(* IEC 61131-3 sources: SortJet_MasterSPS_Aufbau.fbsproj/Device.device.xml.v3^/Plc Logic.plclogic.xml.v3^/Application.application.xml.v3^/09_Station/Stationen/Aufgabe- Anlege- Wand[208]/0_Konfig, 3 files *)

(* ---- Antriebsinformationen_208.gvl ---- *)
(* METADATA
{
	"v3Meta": {
		"objectGuid": "0ee05288-750e-42b2-bc5b-835c7c5d3b07"
	}
}
*)
{attribute 'allow_unqualified_access'}
NAMESPACE Antriebsinformationen_208
VAR_GLOBAL

//-------------------------------------------------------------------------------------------------
// ANTRIEBSINFORMATION
//-------------------------------------------------------------------------------------------------

  apgInfoStation208Glastransport : ARRAY[cWAND_1..cANZAHL_WAENDE] OF AntriebsInformationen := [
    (
      wAchsID                                 :=     15,   // Achs ID aus dem EConSet
      stTyp                                   := 'Belt',  // Typ
      wpSchaltschrank                         :=   2080,  // Daten aus dem Schaltplan
      wpSchaltplanreihe                       :=      2,  // Daten aus dem Schaltplan
      wpSchaltplanseite                       :=    100,  // Daten aus dem Schaltplan
      rpMaxGeschwindigkeit                    :=   1000,  // [mm/s]   Max- Geschwindigkeit für den Automatikbetrieb
      rpHandGeschwindigkeit                   :=    333,  // [mm/s]   Hand- Geschwindigkeit
      rpReduzierteGeschwindigkeit             :=    250,  // [mm/s]   Reduzierte Geschwindigkeit
      rpReferenzGeschwindigkeit               :=     50,  // [mm/s]   Geschwindigkeit für die Referenzfahrt
      rpEinrichtGeschwindigkeit               :=    100,  // [mm/s]   Max Geschwindigkeit während der Einrichtung der Anlage
      rpMaxBeschleunigung                     :=   1500,  // [mm/s^2] Max Beschleunigung
      rpMaxVerzoegerung                       :=   1500,  // [mm/s^2] Max Verzoegerung
      rpMaxRuckzeit                           :=    100,  // [ms]     Ruckzeit des Antriebs
      rpReduzierteBeschleunigung              :=    500,  // [mm/s^2] Reduzierte Beschleunigung
      rpReduzierteVerzoegerung                :=    500,  // [mm/s^2] Reduzierte Verzoegerung
      rpBeschleunigungFremdanlage             :=   1000,  // [mm/s^2] Beschleunigung zu einer Fremdanlage
      rpGeschwindigkeitMessen                 :=    667,  // [mm/s] Geschwindigkeit beim Scheiben messen
      rpGeschwindigkeitSystemcheck            :=  500.0,  // [mm/s]   Geschwindigkeit im Systemcheck (nur Glastransport)
      rpGeschwindigkeitSystemcheckReduzierung :=  167.0,  // [mm/s]   Geschwindigkeit im Systemcheck bei belegtem Vorstop-Sensor (nur Glastransport)
      stOptionen                              := ( eEndschalterQuelle    := Endschalterquelle_EN.KEINE,     // Hardware-Endschalter: KEINE, UMRICHTER oder SPS
                                                   bVersorgungUeberXVR   := FALSE,                          // XVR-Modus: brueckt Hauptschalter 400 V und LS 230 V
                                                   bBremseLoesenFreigabe := FALSE )                         // Der Antrieb darf über eine Betriebsart die Bremse lösen
    )];

  apgInfoStation208GlastransportSlave : ARRAY[cWAND_1..cANZAHL_WAENDE] OF AntriebsInformationen := [
    (
      wAchsID                                 :=     65,   // Achs ID aus dem EConSet
      stTyp                                   := 'Belt',  // Typ
      wpSchaltschrank                         :=   2080,  // Daten aus dem Schaltplan
      wpSchaltplanreihe                       :=      2,  // Daten aus dem Schaltplan
      wpSchaltplanseite                       :=    100,  // Daten aus dem Schaltplan
      rpMaxGeschwindigkeit                    :=   1000,  // [mm/s]   Max- Geschwindigkeit für den Automatikbetrieb
      rpHandGeschwindigkeit                   :=    333,  // [mm/s]   Hand- Geschwindigkeit
      rpReduzierteGeschwindigkeit             :=    250,  // [mm/s]   Reduzierte Geschwindigkeit
      rpReferenzGeschwindigkeit               :=     50,  // [mm/s]   Geschwindigkeit für die Referenzfahrt
      rpEinrichtGeschwindigkeit               :=    100,  // [mm/s]   Max Geschwindigkeit während der Einrichtung der Anlage
      rpMaxBeschleunigung                     :=   1500,  // [mm/s^2] Max Beschleunigung
      rpMaxVerzoegerung                       :=   1500,  // [mm/s^2] Max Verzoegerung
      rpMaxRuckzeit                           :=    100,  // [ms]     Ruckzeit des Antriebs
      rpReduzierteBeschleunigung              :=    500,  // [mm/s^2] Reduzierte Beschleunigung
      rpReduzierteVerzoegerung                :=    500,  // [mm/s^2] Reduzierte Verzoegerung
      rpBeschleunigungFremdanlage             :=   1000,  // [mm/s^2] Beschleunigung zu einer Fremdanlage
      rpGeschwindigkeitMessen                 :=    667,  // [mm/s] Geschwindigkeit beim Scheiben messen
      rpGeschwindigkeitSystemcheck            :=  500.0,  // [mm/s]   Geschwindigkeit im Systemcheck (nur Glastransport)
      rpGeschwindigkeitSystemcheckReduzierung :=  167.0,  // [mm/s]   Geschwindigkeit im Systemcheck bei belegtem Vorstop-Sensor (nur Glastransport)
      stOptionen                              := ( eEndschalterQuelle    := Endschalterquelle_EN.KEINE,     // Hardware-Endschalter: KEINE, UMRICHTER oder SPS
                                                   bVersorgungUeberXVR   := FALSE,                          // XVR-Modus: brueckt Hauptschalter 400 V und LS 230 V
                                                   bBremseLoesenFreigabe := FALSE )                         // Der Antrieb darf über eine Betriebsart die Bremse lösen
    )];

  apgInfoStation208Messachse :  AntriebsInformationen :=
    (
      wAchsID                                 :=        16,   // Achs ID aus dem EConSet
      stTyp                                   := 'Measure',  // Typ
      wpSchaltschrank                         :=      2081,  // Daten aus dem Schaltplan
      wpSchaltplanreihe                       :=         2,  // Daten aus dem Schaltplan
      wpSchaltplanseite                       :=       100,  // Daten aus dem Schaltplan
      rpMaxGeschwindigkeit                    :=      1000,  // [mm/s]   Max- Geschwindigkeit für den Automatikbetrieb
      rpHandGeschwindigkeit                   :=       333,  // [mm/s]   Hand- Geschwindigkeit
      rpReduzierteGeschwindigkeit             :=         0,  // [mm/s]   Reduzierte Geschwindigkeit
      rpReferenzGeschwindigkeit               :=        50,  // [mm/s]   Geschwindigkeit für die Referenzfahrt
      rpEinrichtGeschwindigkeit               :=         0,  // [mm/s]   Max Geschwindigkeit während der Einrichtung der Anlage
      rpMaxBeschleunigung                     :=      2500,  // [mm/s^2] Max Beschleunigung
      rpMaxVerzoegerung                       :=      2500,  // [mm/s^2] Max Verzoegerung
      rpMaxRuckzeit                           :=       500,  // [ms]     Ruckzeit des Antriebs
      rpReduzierteBeschleunigung              :=       500,  // [mm/s^2] Reduzierte Beschleunigung
      rpReduzierteVerzoegerung                :=       500,  // [mm/s^2] Reduzierte Verzoegerung
      rpBeschleunigungFremdanlage             :=         0,  // [mm/s^2] Beschleunigung zu einer Fremdanlage
      rpGeschwindigkeitMessen                 :=         0,  // [mm/s] Geschwindigkeit beim Scheiben messen
      rpGeschwindigkeitSystemcheck            :=     500.0,  // [mm/s]   Geschwindigkeit im Systemcheck (nur Glastransport)
      rpGeschwindigkeitSystemcheckReduzierung :=     167.0,  // [mm/s]   Geschwindigkeit im Systemcheck bei belegtem Vorstop-Sensor (nur Glastransport)
      stOptionen                              := ( eEndschalterQuelle    := Endschalterquelle_EN.UMRICHTER, // Hardware-Endschalter: KEINE, UMRICHTER oder SPS
                                                   bVersorgungUeberXVR   := FALSE,                          // XVR-Modus: brueckt Hauptschalter 400 V und LS 230 V
                                                   bBremseLoesenFreigabe := FALSE )                         // Der Antrieb darf über eine Betriebsart die Bremse lösen
    );

  apgInfoStation208Kippen : AntriebsInformationen :=
    (
      wAchsID                                 :=     65,  // Achs ID aus dem EConSet
      stTyp                                   := 'Tilt',  // Typ
      wpSchaltschrank                         :=      0,  // Daten aus dem Schaltplan
      wpSchaltplanreihe                       :=     02,  // Daten aus dem Schaltplan
      wpSchaltplanseite                       :=      0,  // Daten aus dem Schaltplan
      rpMaxGeschwindigkeit                    :=      0,  // [Grad/s]   Max- Geschwindigkeit für den Automatikbetrieb
      rpHandGeschwindigkeit                   :=      0,  // [Grad/s]   Hand- Geschwindigkeit
      rpReduzierteGeschwindigkeit             :=      0,  // [Grad/s]   Reduzierte Geschwindigkeit
      rpReferenzGeschwindigkeit               :=      0,  // [Grad/s]   Geschwindigkeit für die Referenzfahrt
      rpEinrichtGeschwindigkeit               :=      0,  // [Grad/s]   Max Geschwindigkeit während der Einrichtung der Anlage
      rpMaxBeschleunigung                     :=      0,  // [Grad/s^2] Max Beschleunigung
      rpMaxVerzoegerung                       :=      0,  // [Grad/s^2] Max Verzoegerung
      rpMaxRuckzeit                           :=      0,  // [ms] Ruckzeit des Antriebs
      rpReduzierteBeschleunigung              :=      0,  // [Grad/s^2] Reduzierte Beschleunigung
      rpReduzierteVerzoegerung                :=      0,  // [Grad/s^2] Reduzierte Verzoegerung
      rpBeschleunigungFremdanlage             :=      0,  // [Grad/s^2] Beschleunigung zu einer Fremdanlage
      rpGeschwindigkeitMessen                 :=      0,  // [Grad/s] Geschwindigkeit beim Scheiben messen
      rpGeschwindigkeitSystemcheck            :=  500.0,  // [mm/s]   Geschwindigkeit im Systemcheck (nur Glastransport)
      rpGeschwindigkeitSystemcheckReduzierung :=  167.0,  // [mm/s]   Geschwindigkeit im Systemcheck bei belegtem Vorstop-Sensor (nur Glastransport)
      stOptionen                              := ( eEndschalterQuelle    := Endschalterquelle_EN.KEINE,     // Hardware-Endschalter: KEINE, UMRICHTER oder SPS
                                                   bVersorgungUeberXVR   := FALSE,                          // XVR-Modus: brueckt Hauptschalter 400 V und LS 230 V
                                                   bBremseLoesenFreigabe := FALSE )                         // Der Antrieb darf über eine Betriebsart die Bremse lösen
    );

END_VAR

END_NAMESPACE

(* ---- MK_Station_208.gvl ---- *)
(* METADATA
{
	"v3Meta": {
		"objectGuid": "8432a7e6-a09e-4ecf-ad2f-9f4275e97011"
	}
}
*)
{attribute 'allow_unqualified_access'}
NAMESPACE MK_Station_208
VAR_GLOBAL

//-------------------------------------------------------------------------------------------------
// MASCHINEPARAMETER: ANLEGE- ABNAHME- WAND
//-------------------------------------------------------------------------------------------------

  apgMKStation208 : Parameter_Station :=
    (
      stStationsNummern                     := ( NummerIntern :=  208,                                                       // Stationsnummer fuer das MMI und die Stationsangabe der Meldungen
                                                 NummerExtern := 1208,                                                       // Stationsnummer fuer Bedienermeldungen
                                                 NummerSPS    :=  208                                                        // Stationsnummer SPS-intern (Indizes)
                                               ),
      bDeaktivieren                         := FALSE,                                                                        // Station deaktiviert (keine Auftraege, keine Referenzfahrt)
      wMeldungsNummer                       := 1830,                                                                         // Basis-Meldungsnummer (WatchIO)
      eStationsTyp                          := eStation,                                                                     // Typ der Station
      eaAutomatikkreis                      := [eAutomatikkreis_1],                                                          // Automatikkreise, zu denen die Station gehoert
      eaSicherheitskreis                    := [eSicherheitskreis_Undefiniert],                                              // Sicherheitskreise, in die die Station eingebunden ist
      // astSicherheitskreisTeilabschaltung
      eSystemcheckZyklus                    := eSystemcheckZyklus_1,                                                         // In welchem Zyklus des Systemchecks die Station geprueft wird
      stSchnittstellendaten                 := ( wVorgaengerStation := cSTATION_DEFAULT,                                     // Station vor dieser Station (cSTATION_DYNAMISCH bei mehreren)
                                                 wNachfolgerStation := cSTATION_207,                                         // Station nach dieser Station (cSTATION_DYNAMISCH bei mehreren)
                                                 bStationIstShuttle := FALSE                                                 // Station ist ein Shuttle
                                               ),
      stStationsOptionen                    := ( stSystemcheck :=  ( bScheibenVermessenSystemCheck               := FALSE,   // Scheiben im Systemcheck vermessen
                                                                     bScheibeNachSystemcheckAufAuslauf           := TRUE,    // Scheibe nach dem Systemcheck auf den Auslaufsensor fahren
                                                                     bSystemCheckMitVorgaengerBatchTransport     := FALSE,   // derzeit ohne Funktion
                                                                     bSystemCheckMitNachfolgerBatchTransport     := FALSE,   // derzeit ohne Funktion
                                                                     bOptionSystemCheckScheibeMittigLegen        := FALSE ), // derzeit ohne Funktion

                                                 // stTransfershuttle
                                                 stGlastransport :=  ( bVortransport                             := FALSE,   // Vortransport aktivieren [Bsp.: Nach einem Eintransport mit gesetztem Bit <Letzte Scheibe>]
                                                                       bTransportMasterSlaveEintransport         := FALSE,   // derzeit ohne Funktion
                                                                       bTransportMasterSlaveAustransport         := TRUE ,   // Austransport als Slave auf die Achse des Nachfolgers
                                                                       bGLasUebernahmeSenkrecht                  := FALSE,   // RKT - Eintransport in Senkrechter-Position bzw. in Waagerechter- Position [default]
                                                                       bAustransportISOLinie                     := FALSE,   // Austransport an eine ISO-Linie
                                                                       bScheibenVermessen                        := TRUE,    // Scheibenmessung am Anlegetisch/Anlegewand
                                                                       bMessrichtungNegativ                      := FALSE,   // Negative Fahrtrichtung beim Messen
                                                                       bScheibenmessungEintransport              := FALSE,   // Scheibenmessung beim Eintransport
                                                                       bScheibenmessungSensorVorabAuslauf        := TRUE     // Scheibenmessung mit SensorVorabAuslauf z.B. Anlegewand
                                                                      ),
                                                 stAnlegetisch   :=  ( bIstAnlegestation                         := TRUE,    // Station an der Scheiben angelegt werden [Anlegetisch, Anlegewand]; im Systemcheck-Verbund nur mit genau einer Scheibe
                                                                       bAnschlagAutomatischAusfahren             := FALSE,   // Anschlaege beim Anlegen automatisch ausfahren (Vorgabe, am Taster umschaltbar)
                                                                       bAnlegetischMitEintransportVorgaenger     := FALSE    // VSG: Station entscheidet selbst zwischen Eintransport vom Vorgaenger und Anlegen
                                                                      ),
                                                 // stEckuebergabe
                                                 // stDrehstation
                                                 bVorAbKomponentenAnsteuerung              := FALSE,                         // VorAbKomponentenAnsteuerung Auftraege werden bearbeitet
                                                 bVerstellungEinAusGefahrenLogikDrehen     := FALSE,                         // Verstellung: Logik ein-/ausgefahren gedreht
                                                 bLangsamfahrtNockenQuerfahrtAktivieren    := FALSE,                         // Querfahrt: Langsamfahrt-Nocken auswerten
                                                 bSKBlockierenDurchVorabSensoren           := FALSE,                         // Vorab-Sensoren belegt blockieren das Oeffnen des Sicherheitskreises
                                                 bStationLeerfahrenBeiSkAnforderung        := FALSE,                         // Station bei Anforderung Sicherheitskreis leerfahren
                                                 bScheibeAbnehmenNachEintransport          := TRUE,                          // Scheibe nach dem Eintransport wieder abnehmen
                                                 bGlasAbgenommenAutomatischQuittieren      := FALSE                          // derzeit ohne Funktion
                                               ),
      stStationsAufbau                      := ( bGeblase                      := [ cANZAHL_WAENDE(FALSE) ],                 // Ausbaustufe: Geblaese je Wand
                                                 bGlastransport                := [ TRUE ],                                  // Ausbaustufe: Glastransport je Wand
                                                 bKippen                       := [ cANZAHL_WAENDE(FALSE) ],                 // Ausbaustufe: Kippen je Wand
                                                 bKippenSchuetz                := FALSE,                                     // Kippen ueber Schuetz statt Umrichter
                                                 bTransportVerstellung         := [ cANZAHL_WAENDE(FALSE) ],                 // Ausbaustufe Shuttle: Transport-/Dickenverstellung je Wand
                                                 bHub                          := FALSE,                                     // Ausbaustufe: Hub der Station
                                                 bHubrahmen                    := FALSE,                                     // Ausbaustufe: Hubrahmen (Riemen heben/senken)
                                                 bDrehen                       := FALSE,                                     // Ausbaustufe: Drehen
                                                 bQuerachse                    := FALSE,                                     // Ausbaustufe: Querachse
                                                 bMessachse                    := TRUE,                                      // Ausbaustufe: Messachse (Anlegetisch, Anlegewand)
                                                 bDruckluft                    := FALSE,                                     // Druckluftueberwachung vorhanden
                                                 bAnschlag                     := FALSE,                                     // Ausbaustufe: Ausrichtanschlaege
                                                 bSensorAuslauf                := TRUE,                                      // Auslaufsensor vorhanden
                                                 bSensorEinlauf                := TRUE,                                      // Einlaufsensor vorhanden
                                                 bSensorEinlaufStopp           := FALSE,                                     // Shuttle: zusaetzlicher Stopp-Sensor am Einlauf (ohne: Einlaufsensor), Gegenstueck zum Auslauf-Stopp im Rueckwaertstransport
                                                 bSensorAuslaufStopp           := FALSE,                                     // Shuttle: zusaetzlicher Stopp-Sensor am Auslauf (ohne: Auslaufsensor), Verfahrfreigabe und Scheibe hat Shuttle verlassen
                                                 bDurchlaufSperreZumNachfolger := TRUE,                                      // Ausbaustufe: bewegliche Abschrankung zum Nachfolger
                                                 bQuerfahrt                    := FALSE,                                     // Ausbaustufe: Querfahrt
                                                 bWandverstellung              := [ FALSE ],                                 // Ausbaustufe Station: Wandverstellung je Wand
                                                 bWandverstellungMotorisch     := FALSE,                                     // Shuttle: Transport-/Wandverstellung mit Antrieb statt pneumatisch
                                                 bRoellchenleiste              := [ FALSE ],                                 // Ausbaustufe Station: Roellchenleiste je Wand
                                                 bDurchgang                    := FALSE,                                     // Station ist Teil eines Durchgangs (belegt = Oeffnen blockiert)
                                                 bSlaveAntrieb                 := FALSE,                                     // Glastransport mit Slave-Antrieb
                                                 bRolltor                      := FALSE,                                     // Ausbaustufe Faecherwagen: Rolltor
                                                 bKlemmzylinder                := FALSE,                                     // Ausbaustufe Faecherwagen: Klemmzylinder fixiert den Oberrahmen beim Ein- und Ausschleusen
                                                 bGreifer                      := [cANZAHL_WAENDE(FALSE)],                   // Shuttle: Greifer je Wand (Scheibe aus dem Faecherwagen ziehen bzw. hineinschieben)
                                                 bRFID                         := FALSE,                                     // RFID-Leser vorhanden
                                                 bAGV                          := FALSE,                                     // Ausbaustufe Faecherwagen: Betrieb mit AGV
                                                 bKipparme                     := FALSE,                                     // Ausbaustufe: Kipparme
                                                 bMessachseAmEndeVomTisch      := FALSE,                                     // Messachse am Ende des Tisches (Hoehenfehler fragt den Bediener)
                                                 bDLSSchmiersystem             := FALSE,                                     // Zentralschmierung DLS vorhanden
                                                 bGlastransportSlaveVorhanden  := FALSE,                                     // Glastransport mit Slave-Antrieb (Meldungen/Ueberwachung Slave)
                                                 wHydraulikstation             := 0                                          // Faecherwagen Hydraulik: zugeordnete Hydraulikstation (cHYDRAULIKSTATION_x), 0 = keine
                                               ),
      stStationsParameter                   := ( rLaengeUebergroesseScheibe              := 6000,                            // Shuttle: ab dieser Scheibenlaenge gilt die Scheibe als uebergross [mm]
                                                 rMinGlasHoeheAutomatischenEintransport  := 0.0,                             // VSG: Mindesthoehe fuer automatischen Eintransport [mm]
                                                 rMinGlasLaengeAutomatischenEintransport := 0.0,                             // VSG: Mindestlaenge fuer automatischen Eintransport [mm]
                                                 wMaximaleAnzahlAktiverAuftraege         := 0,                               // derzeit ohne Funktion
                                                 rMinPosSwEsEingrenzung                  := 0.0,                             // Externer zusaetzlicher Software-Endschalter MIN; 0 = inaktiv; darf den MK-MIN nur weiter eingrenzen
                                                 rMaxPosSwEsEingrenzung                  := 0.0,                             // Externer zusaetzlicher Software-Endschalter MAX; 0 = inaktiv; darf den MK-MAX nur weiter eingrenzen
                                                 rPosFreigabePufferAusfahren             := 0.0                              // derzeit ohne Funktion
                                               ),
      // stFremdanlage
      stGlasdaten                           := [( rlMinGlasLaenge := 350,                                                    // minimal zulässige GlasLänge
                                                  rlMaxGlasLaenge := 2500,                                                   // maximale zulässige GlasLänge
                                                  rlMinGlasHoehe  := 190,                                                    // minimal zulässige GlasHöhe
                                                  rlMaxGlasHoehe  := 1800,                                                   // maximale zulässige GlasHöhe
                                                  rlMinGlasDicke  := 3,                                                    // minimal zulässige GlasDicke
                                                  rlMaxGlasDicke  := 12.76,                                                     // maximal zulaessige Glasdicke [mm]
                                                  rlLaengeMaxGlas := 0.0                                                     // maximal zulaessige Glaslaenge [mm]
                                               )]
      // astShuttleAnhaltenQuellen
     );

   apgMKStation208Glastransport : ARRAY[cWAND_1..cANZAHL_WAENDE] OF Parameter_Glastransport := [
    (
      rLaengeStation                        :=  3300, // Länge der Station
      rScheibenabstand                      :=   300, // Der Abstand zwischen zwei Scheiben auf der Station
      rWegUeberAuslauf                      :=    50, // Weg ueber den Auslaufsensor hinaus [mm]
      rWegUeberEinlauf                      :=    50, // Weg ueber den Einlaufsensor hinaus [mm]
      rWegUeberSensorenSystemCheck          :=    15, // Der Weg der Ueber ein die Sensoren zum vermessen der Scheiben
      rUeberwachungAuslaufsensor            :=   500, // Ueberwachung des Auslaufsensors [Strecke in der der Auslaufsensor Frei / ueberfahren werden soll]
      rUeberwachungEinlaufsensor            :=   500, // Ueberwachung des Einlaufsensors [Strecke in der der Einlaufsensor Frei / ueberfahren werden soll]
      rWegUeberEinlaufEintransport          :=    30, // Eintransport vorwaerts: Abstand Scheibenhinterkante zum Einlaufsensor [mm]
      rWegUeberEinlaufAustransport          :=    30, // Lage Auf Einlauf: Scheibe liegt um diesen Weg auf dem Einlaufsensor [mm]
      rWegUeberAuslaufEintransport          :=    30, // Eintransport rueckwaerts: Abstand Scheibenhinterkante zum Auslaufsensor [mm]
      rWegUeberAuslaufAustransport          :=    15, // Lage Auf Auslauf: Weg ueber den Auslaufsensor hinaus [mm]
      rWegEinlaufsensorZuVorStopSensor      :=  3160, // Beschreibt den Weg vum eine Scheibe beim EIntransport vom Einlaufsensor bis ueberden Vorabstopsensor zu verfahren
      rMesstoleranz                         :=    10, // Toleranz-Mass fuer die Scheibenlaengenmessung
      rMessstrecke                          :=  2904, // Beschreibt die Strecke ziwischen 2 Sensoren die der Antrieb verfaehrt
      rWegstreckeBisZurVerzoegerung         :=  2660  // Beschreibt die Strecke die gefahren werden soll bis der Antrieb abgebremst werden soll, dies gilt fuer Eintransportauftraege die das Bit "Letzte Scheibe" gesetzt haben
    )];

  apgMKStation208Messachse: Parameter_Messachse :=
    (
      rKorrekturOffset                      :=    0, // Korrektur der Position um einen Bestimmten Wert (Offset)
      rStreckePositionieren                 :=    0, // ?
      rPositionUeberScheibenhoehe           := 0.0,  // Position der Zentrierleiste ueber dem Glas so dass das Glas angelegt werden kann
      rVerfahrbereichsOffset                := 0.0,  // Korrektur des Verfahrens wenn
      rKorrekturOffsetVSGEintransport       := 0.0,  // Korrektur der Position um einen Bestimmten Wert (Offset) beim Eintransport von VSG
      rOffsetMessung                        := 0.0,  // ?
      rToleranz                             := 0.0,  // Toleranzwert in der Ausmessung der Höhe
      rAbstandSensorenOberUndUnterkante     := 0.0,  // Rechnerischer Abstand zwischen dem Sensor der die Scheibenunterkante misst und dem Sensor der die Scheibenoberkante misst
      rOffsetNullLinie                      := 0.0   // Offset das auf den Wert des Abstands zur Null-Linie aufgerechnet wird, um dies evtl zu korrigieren
    );

  apgMKStation208Kippen : ARRAY[cWAND_1..cANZAHL_WAENDE] OF Parameter_Kippen := [
    (
      tZeitlicheUeberwachungKippen          := TIME#5000MS, // [ms \ s] Verwendet fuer Antriebe die Ueber einen Schuetz angesteuert werden
      tZeitAntriebsfreigabeErhalten         :=  TIME#180S,  // [ms \ s] Energieeinsparrung: Zeiteinheit nach der die Antriebsfreigabe entzogen werden soll wenn keine Aktion ansteht [1 s = 1000 ms ]
      rToleranz                             :=          1,  // Toleranz beim Entscheiden der aktuellen Position
      rPosition0Grad                        :=          0,  // Waagerechte- Position 0 Grad: Position auf die die Station gehoben werden soll
      rPosition90Grad                       :=          0,  // Senkrechte-Position 90 Grad : Position auf die die Station gesenkt werden soll
      bKippenMitSchuetz                     :=      FALSE,  // Kippen per Umrichter oder Schütz
      rPosition84Grad                       := 0.0,         // Senkrechte- Position 84 Grad: Position auf die die Station gehoben werden soll
      rPosition88_5Grad                     := 0.0,         // Senkrechte- Position 84 Grad: Position auf die die Station gehoben werden soll
      rPosition96Grad                       := 0.0          // Senkrechte-Position 96 Grad : Position auf die die Station gesenkt werden soll
    )];

END_VAR
END_NAMESPACE

(* ---- Konfiguration_208.gvl ---- *)
(* METADATA
{
	"v3Meta": {
		"objectGuid": "94633f29-785d-43e8-8fe9-544c355e9fea"
	}
}
*)
{attribute 'allow_unqualified_access'}
NAMESPACE Konfiguration_208
VAR_CONFIG

  // Taster
  Globale_Bausteine.Combiwand208.in_bFussTasterGlasAngelegt                               AT %MX1.0    : BOOL; // OPTION - Signal Scheibe ist angelegt Fusstaster
  Globale_Bausteine.Combiwand208.in_bTasterGlasAngelegt                                   AT %IX3.7    : BOOL; // IO-L - 208 quittieren Scheibe aufgelegt
  Globale_Bausteine.Combiwand208.in_bTasterFehlmessungQuittiern                           AT %IX4.0    : BOOL; // IO-L - 208 Fehlmessung quittieren
  Globale_Bausteine.Combiwand208.in_bKnebelGlastransportZurueck                           AT %IX4.2    : BOOL; // IO-L - 208 Riemen zurueck
  Globale_Bausteine.Combiwand208.in_bKnebelGlastransportVor                               AT %IX4.1    : BOOL; // IO-L - 208 Riemen vor
  Globale_Bausteine.Combiwand208.in_bTasterGlasbruch                                      AT %IX4.3    : BOOL; // IO-L - 208 Glasbruch
  Globale_Bausteine.Combiwand208.in_bTasterQuittierungGlasAbgenommen                      AT %IX3.7    : BOOL; // IO-L - 208 quittieren Scheibe aufgelegt (gleicher Taster wie Glas angelegt)

  // Lampen/Ampel
  Globale_Bausteine.Combiwand208.out_bAmpelSignalGruen                                    AT %QX5.0    : BOOL; // IO-L - 208 Freigabe Scheibe anlegen Ampel gruen
  Globale_Bausteine.Combiwand208.out_bSignalScheibeAufgegeben                             AT %QX4.5    : BOOL; // IO-L - 208 quittieren Scheibe aufgelegt
  Globale_Bausteine.Combiwand208.out_bSignalScheibeFehlmessung                            AT %QX4.6    : BOOL; // IO-L - 208 Scheibe Fehlmessung
  Globale_Bausteine.Combiwand208.out_bSignalScheibeGlasbruch                              AT %QX4.7    : BOOL; // IO-L - 208 Glasbruch Meldung
  Globale_Bausteine.Combiwand208.out_bSignalScheibeAbnehmen                               AT %MX2080.1 : BOOL; // OPTION

  // Bewegliche Abschrankung zum Nachfolger (geschlossen kommt ueber die Safety)
  Globale_Bausteine.Combiwand208.in_bSensorAbschrankungOffen                              AT %IX9.0    : BOOL; // IO-L - 208 bewegliche Abschrankung offen
  Globale_Bausteine.Combiwand208.out_bAbschrankungEinfahren                               AT %QX10.4   : BOOL; // IO-L - 208 bewegliche Abschrankung einfahren (oeffnen)
  Globale_Bausteine.Combiwand208.out_bAbschrankungAusfahren                               AT %QX10.5   : BOOL; // IO-L - 208 bewegliche Abschrankung ausfahren (schliessen)

  // Lichtschranke
  Globale_Bausteine.Combiwand208.in_bLichtschrankeQuittiert                               AT %MX1.1    : BOOL; // OPTION
  Globale_Bausteine.Combiwand208.in_bLichtschrankeFehler                                  AT %MX1.1    : BOOL; // OPTION
  Globale_Bausteine.Combiwand208.out_bLichtschrankeAusgeloest                             AT %MX2080.2 : BOOL; // OPTION - Lichtschranke an der Station ausgelöst und nicht quittiert

  // Gebläse
  Globale_Bausteine.Combiwand208.in_bTasterGeblaeseEin                                    AT %MX1.0     : BOOL; // OPTION - Taster Geblaese ein
  Globale_Bausteine.Combiwand208.in_bMotorschutzGeblaese_Ok                               AT %MX1.1     : BOOL; // OPTION - Motorschutzschalter / Sicherung des Antriebs
  Globale_Bausteine.Combiwand208.out_bGeblaeseEin                                         AT %MX2080.3  : BOOL; // OPTION - Geblaese starten (Schuetz)

  // Dickenverstellung
  Globale_Bausteine.Combiwand208.Dickenverstellung.in_bStatusZylinder1Ausgefahren         AT %MX1.0     : BOOL; // OPTION
  Globale_Bausteine.Combiwand208.Dickenverstellung.in_bStatusZylinder1Eingefahren         AT %MX1.0     : BOOL; // OPTION
  Globale_Bausteine.Combiwand208.Dickenverstellung.in_bStatusZylinder2Ausgefahren         AT %MX1.0     : BOOL; // OPTION
  Globale_Bausteine.Combiwand208.Dickenverstellung.in_bStatusZylinder2Eingefahren         AT %MX1.0     : BOOL; // OPTION

  Globale_Bausteine.Combiwand208.Dickenverstellung.out_bZylinder1Ausfahren                AT %MX2080.4  : BOOL; // OPTION
  Globale_Bausteine.Combiwand208.Dickenverstellung.out_bZylinder1Einfahren                AT %MX2080.5  : BOOL; // OPTION
  Globale_Bausteine.Combiwand208.Dickenverstellung.out_bZylinder2Ausfahren                AT %MX2080.6  : BOOL; // OPTION
  Globale_Bausteine.Combiwand208.Dickenverstellung.out_bZylinder2Einfahren                AT %MX2080.7  : BOOL; // OPTION

  // Kippen
  Globale_Bausteine.Combiwand208.Kippen.in_bMotorschutzschalter_OK                        AT %MX1.1     : BOOL; // OPTION
  Globale_Bausteine.Combiwand208.Kippen.in_bMotorstarter_OK                               AT %MX1.1     : BOOL; // OPTION
  Globale_Bausteine.Combiwand208.Kippen.in_bLSBremse_OK                                   AT %MX1.1     : BOOL; // OPTION
  Globale_Bausteine.Combiwand208.Kippen.in_bLS400V_OK                                     AT %MX1.1     : BOOL; // OPTION

  Globale_Bausteine.Combiwand208.Kippen.out_bKippen84Grad                                 AT %MX2081.0  : BOOL; // OPTION
  Globale_Bausteine.Combiwand208.Kippen.out_bKippen90Grad                                 AT %MX2081.1  : BOOL; // OPTION
  Globale_Bausteine.Combiwand208.Kippen.out_bBremseLoesen                                 AT %MX2081.2  : BOOL; // OPTION
  Globale_Bausteine.Combiwand208.Kippen.out_bReset                                        AT %MX2081.3  : BOOL; // OPTION

  // Nicht vorhandene Komponenten (der Basic erwartet sie, die Instanzen bleiben deaktiviert): Eingaenge auf %MX1.x, Ausgaenge auf freie Merker

  // Hub (unbenutzt)
  Globale_Bausteine.Combiwand208.HubUnbenutzt.in_bSensorNichtUnten                                AT %MX1.0   : BOOL; // OPTION
  Globale_Bausteine.Combiwand208.HubUnbenutzt.in_bSensorNichtOben                                 AT %MX1.0   : BOOL; // OPTION
  Globale_Bausteine.Combiwand208.HubUnbenutzt.in_bMotorstarter_OK                                 AT %MX1.1   : BOOL; // OPTION
  Globale_Bausteine.Combiwand208.HubUnbenutzt.in_bLSBremse_OK                                     AT %MX1.1   : BOOL; // OPTION
  Globale_Bausteine.Combiwand208.HubUnbenutzt.in_bLS400V_OK                                       AT %MX1.1   : BOOL; // OPTION
  Globale_Bausteine.Combiwand208.HubUnbenutzt.out_bHubAbSetzen                                    AT %MX2081.4 : BOOL; // OPTION
  Globale_Bausteine.Combiwand208.HubUnbenutzt.out_bHubAufSetzen                                   AT %MX2081.5 : BOOL; // OPTION
  Globale_Bausteine.Combiwand208.HubUnbenutzt.out_bReset                                          AT %MX2081.6 : BOOL; // OPTION
  Globale_Bausteine.Combiwand208.HubUnbenutzt.out_bBremseLoesen                                   AT %MX2081.7 : BOOL; // OPTION

  // Roellchenleiste (unbenutzt)
  Globale_Bausteine.Combiwand208.RoellchenleisteUnbenutzt.in_bStatusZylinder1Ausgefahren          AT %MX1.0   : BOOL; // OPTION
  Globale_Bausteine.Combiwand208.RoellchenleisteUnbenutzt.in_bStatusZylinder1Eingefahren          AT %MX1.0   : BOOL; // OPTION
  Globale_Bausteine.Combiwand208.RoellchenleisteUnbenutzt.in_bStatusZylinder2Ausgefahren          AT %MX1.0   : BOOL; // OPTION
  Globale_Bausteine.Combiwand208.RoellchenleisteUnbenutzt.in_bStatusZylinder2Eingefahren          AT %MX1.0   : BOOL; // OPTION
  Globale_Bausteine.Combiwand208.RoellchenleisteUnbenutzt.out_bZylinder1Ausfahren                 AT %MX2082.0 : BOOL; // OPTION
  Globale_Bausteine.Combiwand208.RoellchenleisteUnbenutzt.out_bZylinder1Einfahren                 AT %MX2082.1 : BOOL; // OPTION
  Globale_Bausteine.Combiwand208.RoellchenleisteUnbenutzt.out_bZylinder2Ausfahren                 AT %MX2082.2 : BOOL; // OPTION
  Globale_Bausteine.Combiwand208.RoellchenleisteUnbenutzt.out_bZylinder2Einfahren                 AT %MX2082.3 : BOOL; // OPTION

  // Wandverstellung (unbenutzt)
  Globale_Bausteine.Combiwand208.WandverstellungUnbenutzt.in_bStatusZylinder1Ausgefahren          AT %MX1.0   : BOOL; // OPTION
  Globale_Bausteine.Combiwand208.WandverstellungUnbenutzt.in_bStatusZylinder1Eingefahren          AT %MX1.0   : BOOL; // OPTION
  Globale_Bausteine.Combiwand208.WandverstellungUnbenutzt.in_bStatusZylinder2Ausgefahren          AT %MX1.0   : BOOL; // OPTION
  Globale_Bausteine.Combiwand208.WandverstellungUnbenutzt.in_bStatusZylinder2Eingefahren          AT %MX1.0   : BOOL; // OPTION
  Globale_Bausteine.Combiwand208.WandverstellungUnbenutzt.out_bZylinder1Ausfahren                 AT %MX2082.4 : BOOL; // OPTION
  Globale_Bausteine.Combiwand208.WandverstellungUnbenutzt.out_bZylinder1Einfahren                 AT %MX2082.5 : BOOL; // OPTION
  Globale_Bausteine.Combiwand208.WandverstellungUnbenutzt.out_bZylinder2Ausfahren                 AT %MX2082.6 : BOOL; // OPTION
  Globale_Bausteine.Combiwand208.WandverstellungUnbenutzt.out_bZylinder2Einfahren                 AT %MX2082.7 : BOOL; // OPTION

  // Geblaese-Baustein (Motorschutz und Ausgang kommen von der Station)
  Globale_Bausteine.Combiwand208.Geblaese.in_bMotorschutzschalter_OK                     AT %MX1.1   : BOOL; // OPTION
  Globale_Bausteine.Combiwand208.Geblaese.out_bStarteGeblaese                            AT %MX2083.0 : BOOL; // OPTION

END_VAR
END_NAMESPACE
